Fanuc KAREL source: KA00219.KL

PROGRAM KA00219
%NOLOCKGROUP
VAR
  SRC: ARRAY[4] OF JOINTPOS
  DST: ARRAY[4] OF BOOLEAN
BEGIN
  DST = SRC
END KA00219
